(* Logix 5000 project; controller CIP vendor 1 type 14 code 106 rev 20.12; software revision 20.06; part 9 of 13 *)
(* tags used below, declared in another part *)
   MOA_OFF : DINT[10];
   MOA_ON : DINT[10];
   PV_Output_Status : INT[10];
   PV_Output_Status_IND : INT[10,16];
   PV_Status_Bit : BOOL;
(* MainProgram, continued *)

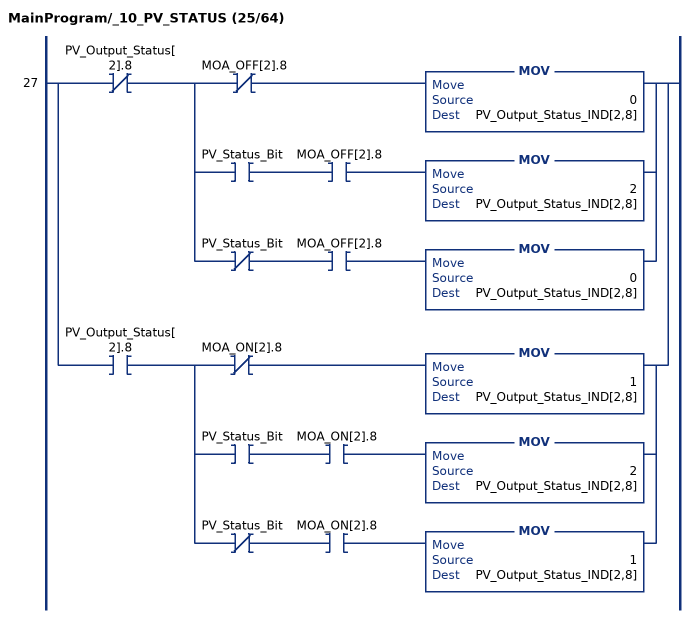
   [picture p157: MainProgram/_10_PV_STATUS rungs 27-27]
   27: [XIO(PV_Output_Status[2].8) [XIO(MOA_OFF[2].8) MOV(0,PV_Output_Status_IND[2,8]) ,XIC(PV_Status_Bit) XIC(MOA_OFF[2].8) MOV(2,PV_Output_Status_IND[2,8]) ,XIO(PV_Status_Bit) XIC(MOA_OFF[2].8) MOV(0,PV_Output_Status_IND[2,8]) ] ,XIC(PV_Output_Status[2].8) [XIO(MOA_ON[2].8) MOV(1,PV_Output_Status_IND[2,8]) ,XIC(PV_Status_Bit) XIC(MOA_ON[2].8) MOV(2,PV_Output_Status_IND[2,8]) ,XIO(PV_Status_Bit) XIC(MOA_ON[2].8) MOV(1,PV_Output_Status_IND[2,8]) ] ];
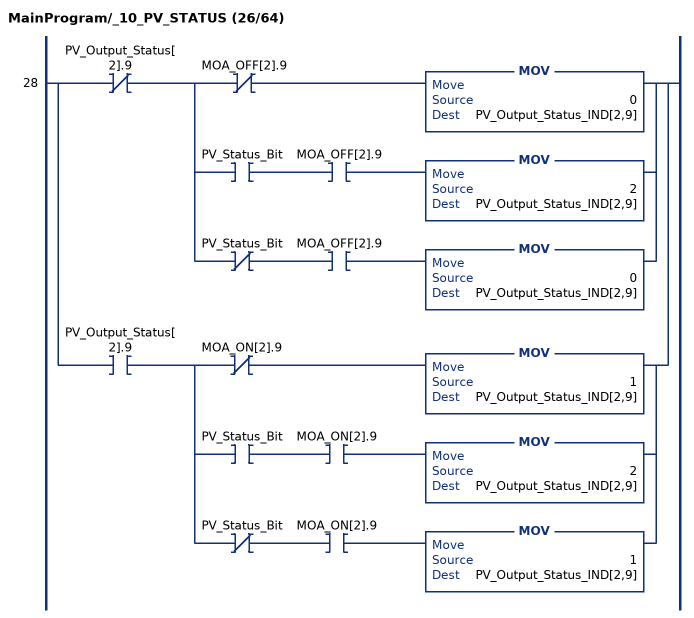
   28: [XIO(PV_Output_Status[2].9) [XIO(MOA_OFF[2].9) MOV(0,PV_Output_Status_IND[2,9]) ,XIC(PV_Status_Bit) XIC(MOA_OFF[2].9) MOV(2,PV_Output_Status_IND[2,9]) ,XIO(PV_Status_Bit) XIC(MOA_OFF[2].9) MOV(0,PV_Output_Status_IND[2,9]) ] ,XIC(PV_Output_Status[2].9) [XIO(MOA_ON[2].9) MOV(1,PV_Output_Status_IND[2,9]) ,XIC(PV_Status_Bit) XIC(MOA_ON[2].9) MOV(2,PV_Output_Status_IND[2,9]) ,XIO(PV_Status_Bit) XIC(MOA_ON[2].9) MOV(1,PV_Output_Status_IND[2,9]) ] ];
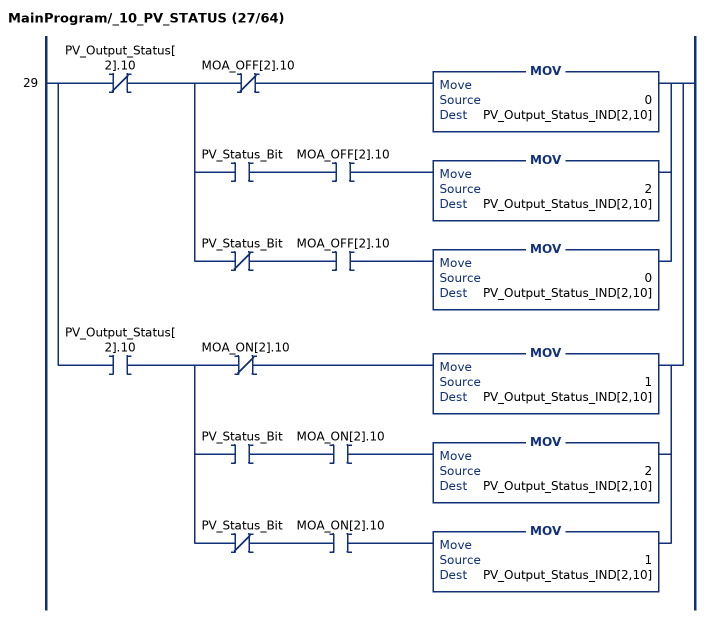
   29: [XIO(PV_Output_Status[2].10) [XIO(MOA_OFF[2].10) MOV(0,PV_Output_Status_IND[2,10]) ,XIC(PV_Status_Bit) XIC(MOA_OFF[2].10) MOV(2,PV_Output_Status_IND[2,10]) ,XIO(PV_Status_Bit) XIC(MOA_OFF[2].10) MOV(0,PV_Output_Status_IND[2,10]) ] ,XIC(PV_Output_Status[2].10) [XIO(MOA_ON[2].10) MOV(1,PV_Output_Status_IND[2,10]) ,XIC(PV_Status_Bit) XIC(MOA_ON[2].10) MOV(2,PV_Output_Status_IND[2,10]) ,XIO(PV_Status_Bit) XIC(MOA_ON[2].10) MOV(1,PV_Output_Status_IND[2,10]) ] ];
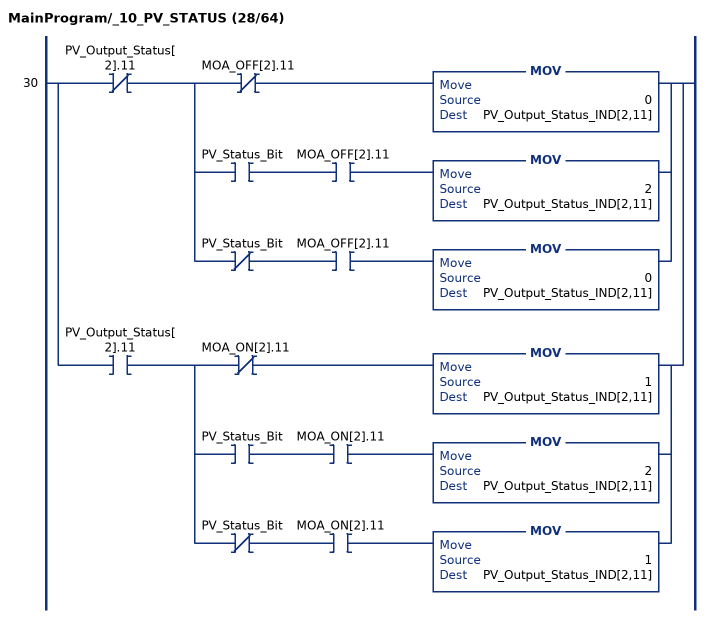
   30: [XIO(PV_Output_Status[2].11) [XIO(MOA_OFF[2].11) MOV(0,PV_Output_Status_IND[2,11]) ,XIC(PV_Status_Bit) XIC(MOA_OFF[2].11) MOV(2,PV_Output_Status_IND[2,11]) ,XIO(PV_Status_Bit) XIC(MOA_OFF[2].11) MOV(0,PV_Output_Status_IND[2,11]) ] ,XIC(PV_Output_Status[2].11) [XIO(MOA_ON[2].11) MOV(1,PV_Output_Status_IND[2,11]) ,XIC(PV_Status_Bit) XIC(MOA_ON[2].11) MOV(2,PV_Output_Status_IND[2,11]) ,XIO(PV_Status_Bit) XIC(MOA_ON[2].11) MOV(1,PV_Output_Status_IND[2,11]) ] ];
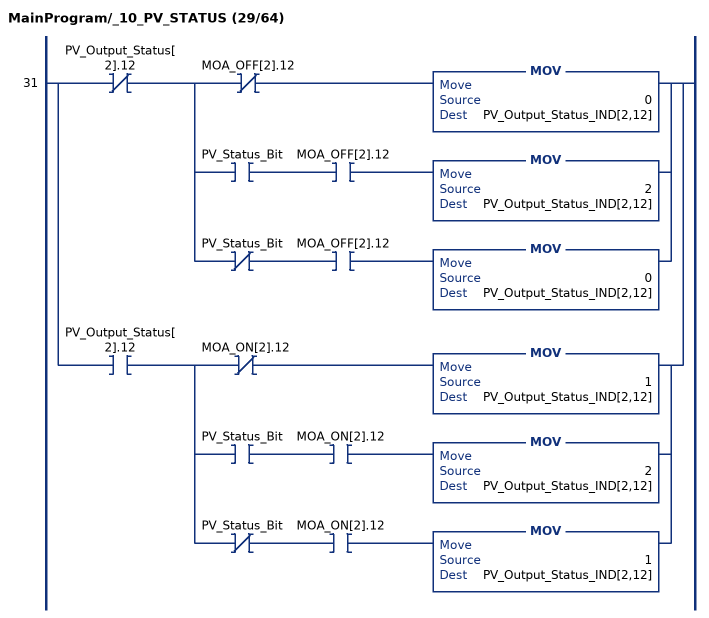
   31: [XIO(PV_Output_Status[2].12) [XIO(MOA_OFF[2].12) MOV(0,PV_Output_Status_IND[2,12]) ,XIC(PV_Status_Bit) XIC(MOA_OFF[2].12) MOV(2,PV_Output_Status_IND[2,12]) ,XIO(PV_Status_Bit) XIC(MOA_OFF[2].12) MOV(0,PV_Output_Status_IND[2,12]) ] ,XIC(PV_Output_Status[2].12) [XIO(MOA_ON[2].12) MOV(1,PV_Output_Status_IND[2,12]) ,XIC(PV_Status_Bit) XIC(MOA_ON[2].12) MOV(2,PV_Output_Status_IND[2,12]) ,XIO(PV_Status_Bit) XIC(MOA_ON[2].12) MOV(1,PV_Output_Status_IND[2,12]) ] ];
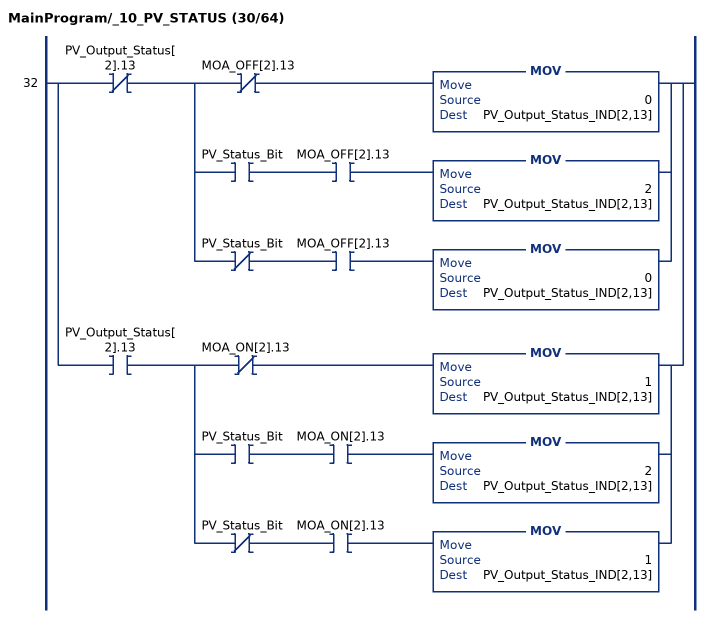
   32: [XIO(PV_Output_Status[2].13) [XIO(MOA_OFF[2].13) MOV(0,PV_Output_Status_IND[2,13]) ,XIC(PV_Status_Bit) XIC(MOA_OFF[2].13) MOV(2,PV_Output_Status_IND[2,13]) ,XIO(PV_Status_Bit) XIC(MOA_OFF[2].13) MOV(0,PV_Output_Status_IND[2,13]) ] ,XIC(PV_Output_Status[2].13) [XIO(MOA_ON[2].13) MOV(1,PV_Output_Status_IND[2,13]) ,XIC(PV_Status_Bit) XIC(MOA_ON[2].13) MOV(2,PV_Output_Status_IND[2,13]) ,XIO(PV_Status_Bit) XIC(MOA_ON[2].13) MOV(1,PV_Output_Status_IND[2,13]) ] ];
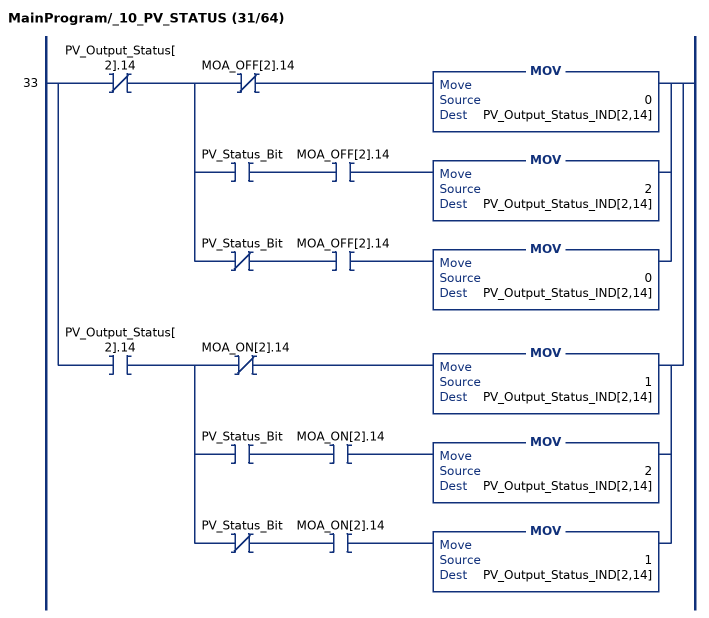
   33: [XIO(PV_Output_Status[2].14) [XIO(MOA_OFF[2].14) MOV(0,PV_Output_Status_IND[2,14]) ,XIC(PV_Status_Bit) XIC(MOA_OFF[2].14) MOV(2,PV_Output_Status_IND[2,14]) ,XIO(PV_Status_Bit) XIC(MOA_OFF[2].14) MOV(0,PV_Output_Status_IND[2,14]) ] ,XIC(PV_Output_Status[2].14) [XIO(MOA_ON[2].14) MOV(1,PV_Output_Status_IND[2,14]) ,XIC(PV_Status_Bit) XIC(MOA_ON[2].14) MOV(2,PV_Output_Status_IND[2,14]) ,XIO(PV_Status_Bit) XIC(MOA_ON[2].14) MOV(1,PV_Output_Status_IND[2,14]) ] ];
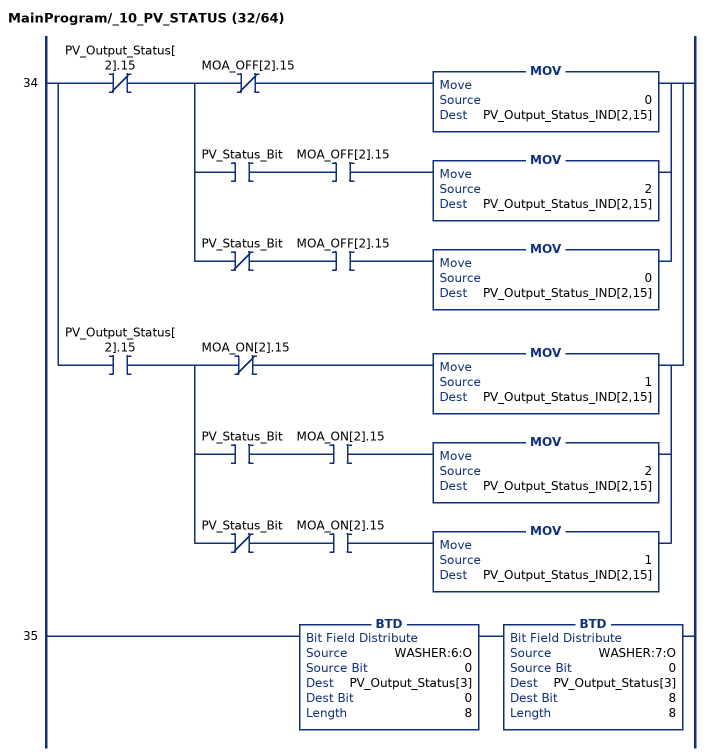
   34: [XIO(PV_Output_Status[2].15) [XIO(MOA_OFF[2].15) MOV(0,PV_Output_Status_IND[2,15]) ,XIC(PV_Status_Bit) XIC(MOA_OFF[2].15) MOV(2,PV_Output_Status_IND[2,15]) ,XIO(PV_Status_Bit) XIC(MOA_OFF[2].15) MOV(0,PV_Output_Status_IND[2,15]) ] ,XIC(PV_Output_Status[2].15) [XIO(MOA_ON[2].15) MOV(1,PV_Output_Status_IND[2,15]) ,XIC(PV_Status_Bit) XIC(MOA_ON[2].15) MOV(2,PV_Output_Status_IND[2,15]) ,XIO(PV_Status_Bit) XIC(MOA_ON[2].15) MOV(1,PV_Output_Status_IND[2,15]) ] ];
   35: BTD(WASHER:6:O,0,PV_Output_Status[3],0,8)BTD(WASHER:7:O,0,PV_Output_Status[3],8,8);
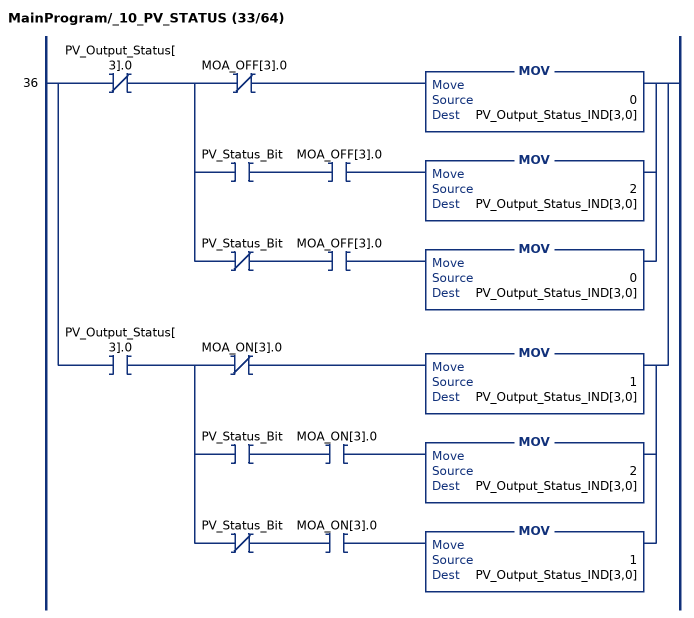
   36: [XIO(PV_Output_Status[3].0) [XIO(MOA_OFF[3].0) MOV(0,PV_Output_Status_IND[3,0]) ,XIC(PV_Status_Bit) XIC(MOA_OFF[3].0) MOV(2,PV_Output_Status_IND[3,0]) ,XIO(PV_Status_Bit) XIC(MOA_OFF[3].0) MOV(0,PV_Output_Status_IND[3,0]) ] ,XIC(PV_Output_Status[3].0) [XIO(MOA_ON[3].0) MOV(1,PV_Output_Status_IND[3,0]) ,XIC(PV_Status_Bit) XIC(MOA_ON[3].0) MOV(2,PV_Output_Status_IND[3,0]) ,XIO(PV_Status_Bit) XIC(MOA_ON[3].0) MOV(1,PV_Output_Status_IND[3,0]) ] ];
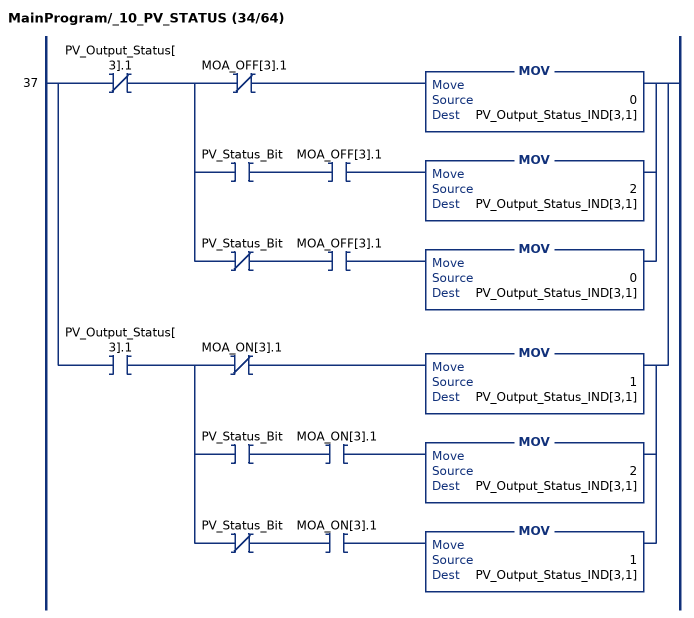
   37: [XIO(PV_Output_Status[3].1) [XIO(MOA_OFF[3].1) MOV(0,PV_Output_Status_IND[3,1]) ,XIC(PV_Status_Bit) XIC(MOA_OFF[3].1) MOV(2,PV_Output_Status_IND[3,1]) ,XIO(PV_Status_Bit) XIC(MOA_OFF[3].1) MOV(0,PV_Output_Status_IND[3,1]) ] ,XIC(PV_Output_Status[3].1) [XIO(MOA_ON[3].1) MOV(1,PV_Output_Status_IND[3,1]) ,XIC(PV_Status_Bit) XIC(MOA_ON[3].1) MOV(2,PV_Output_Status_IND[3,1]) ,XIO(PV_Status_Bit) XIC(MOA_ON[3].1) MOV(1,PV_Output_Status_IND[3,1]) ] ];
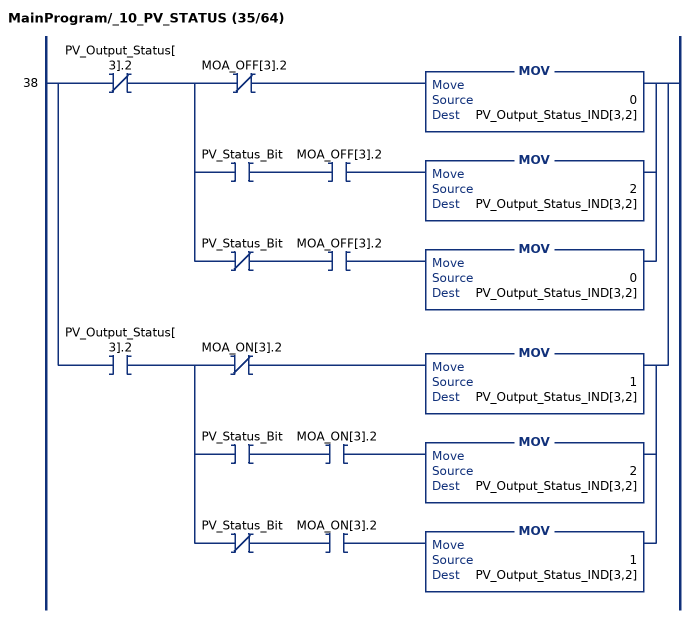
   38: [XIO(PV_Output_Status[3].2) [XIO(MOA_OFF[3].2) MOV(0,PV_Output_Status_IND[3,2]) ,XIC(PV_Status_Bit) XIC(MOA_OFF[3].2) MOV(2,PV_Output_Status_IND[3,2]) ,XIO(PV_Status_Bit) XIC(MOA_OFF[3].2) MOV(0,PV_Output_Status_IND[3,2]) ] ,XIC(PV_Output_Status[3].2) [XIO(MOA_ON[3].2) MOV(1,PV_Output_Status_IND[3,2]) ,XIC(PV_Status_Bit) XIC(MOA_ON[3].2) MOV(2,PV_Output_Status_IND[3,2]) ,XIO(PV_Status_Bit) XIC(MOA_ON[3].2) MOV(1,PV_Output_Status_IND[3,2]) ] ];
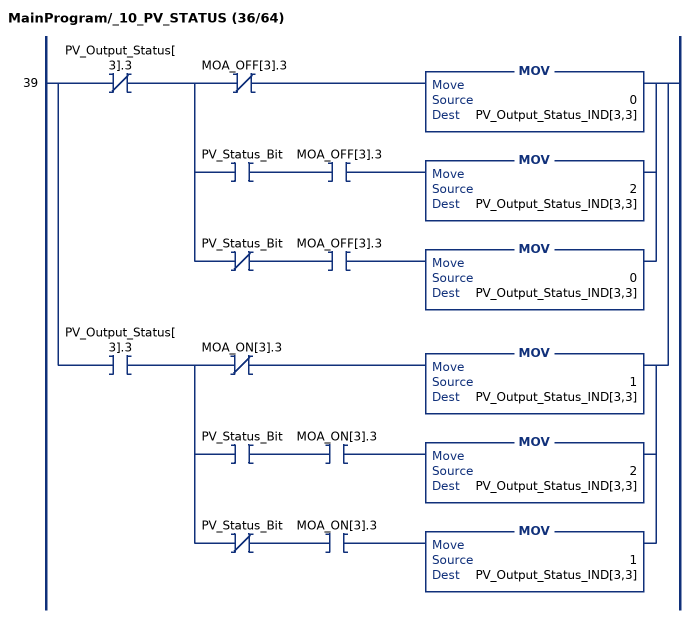
   39: [XIO(PV_Output_Status[3].3) [XIO(MOA_OFF[3].3) MOV(0,PV_Output_Status_IND[3,3]) ,XIC(PV_Status_Bit) XIC(MOA_OFF[3].3) MOV(2,PV_Output_Status_IND[3,3]) ,XIO(PV_Status_Bit) XIC(MOA_OFF[3].3) MOV(0,PV_Output_Status_IND[3,3]) ] ,XIC(PV_Output_Status[3].3) [XIO(MOA_ON[3].3) MOV(1,PV_Output_Status_IND[3,3]) ,XIC(PV_Status_Bit) XIC(MOA_ON[3].3) MOV(2,PV_Output_Status_IND[3,3]) ,XIO(PV_Status_Bit) XIC(MOA_ON[3].3) MOV(1,PV_Output_Status_IND[3,3]) ] ];
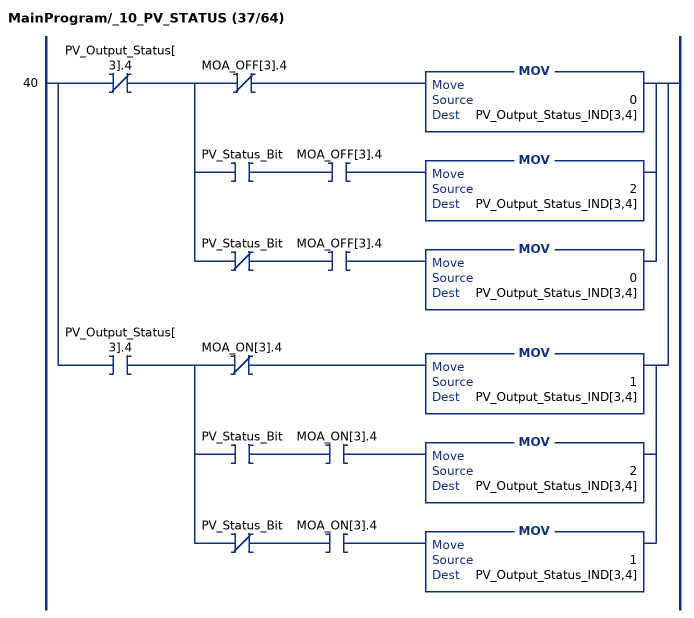
   40: [XIO(PV_Output_Status[3].4) [XIO(MOA_OFF[3].4) MOV(0,PV_Output_Status_IND[3,4]) ,XIC(PV_Status_Bit) XIC(MOA_OFF[3].4) MOV(2,PV_Output_Status_IND[3,4]) ,XIO(PV_Status_Bit) XIC(MOA_OFF[3].4) MOV(0,PV_Output_Status_IND[3,4]) ] ,XIC(PV_Output_Status[3].4) [XIO(MOA_ON[3].4) MOV(1,PV_Output_Status_IND[3,4]) ,XIC(PV_Status_Bit) XIC(MOA_ON[3].4) MOV(2,PV_Output_Status_IND[3,4]) ,XIO(PV_Status_Bit) XIC(MOA_ON[3].4) MOV(1,PV_Output_Status_IND[3,4]) ] ];
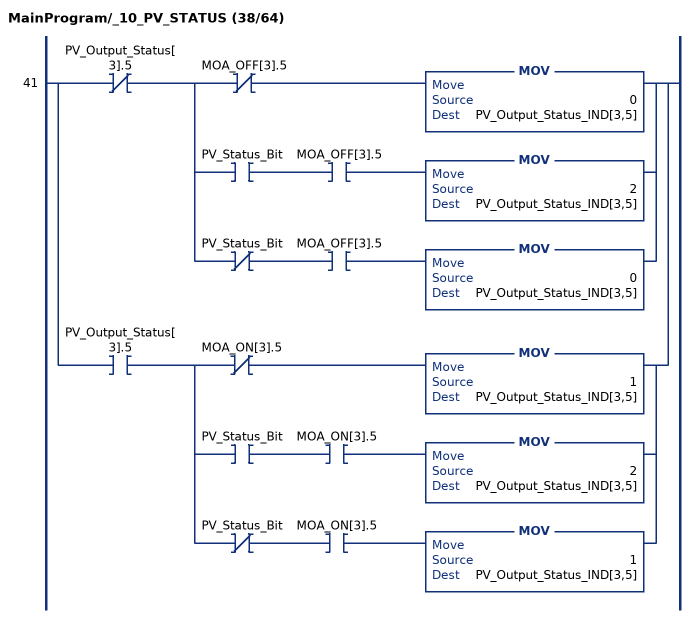
   41: [XIO(PV_Output_Status[3].5) [XIO(MOA_OFF[3].5) MOV(0,PV_Output_Status_IND[3,5]) ,XIC(PV_Status_Bit) XIC(MOA_OFF[3].5) MOV(2,PV_Output_Status_IND[3,5]) ,XIO(PV_Status_Bit) XIC(MOA_OFF[3].5) MOV(0,PV_Output_Status_IND[3,5]) ] ,XIC(PV_Output_Status[3].5) [XIO(MOA_ON[3].5) MOV(1,PV_Output_Status_IND[3,5]) ,XIC(PV_Status_Bit) XIC(MOA_ON[3].5) MOV(2,PV_Output_Status_IND[3,5]) ,XIO(PV_Status_Bit) XIC(MOA_ON[3].5) MOV(1,PV_Output_Status_IND[3,5]) ] ];
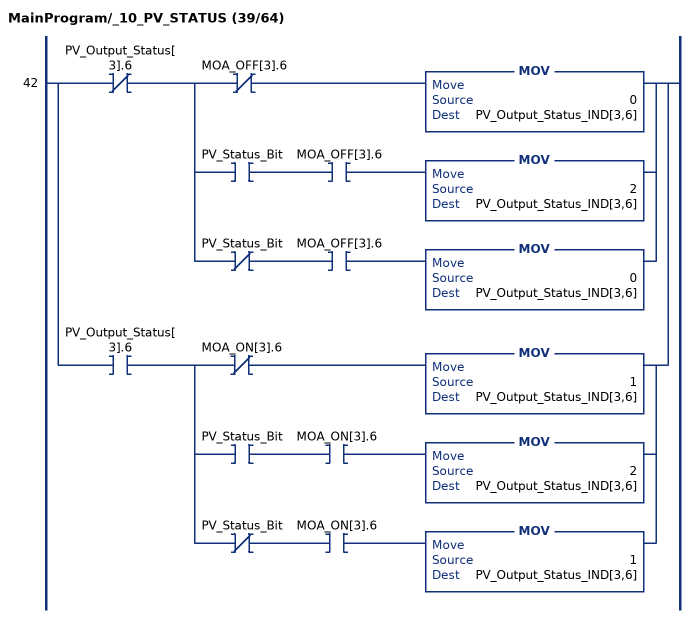
   42: [XIO(PV_Output_Status[3].6) [XIO(MOA_OFF[3].6) MOV(0,PV_Output_Status_IND[3,6]) ,XIC(PV_Status_Bit) XIC(MOA_OFF[3].6) MOV(2,PV_Output_Status_IND[3,6]) ,XIO(PV_Status_Bit) XIC(MOA_OFF[3].6) MOV(0,PV_Output_Status_IND[3,6]) ] ,XIC(PV_Output_Status[3].6) [XIO(MOA_ON[3].6) MOV(1,PV_Output_Status_IND[3,6]) ,XIC(PV_Status_Bit) XIC(MOA_ON[3].6) MOV(2,PV_Output_Status_IND[3,6]) ,XIO(PV_Status_Bit) XIC(MOA_ON[3].6) MOV(1,PV_Output_Status_IND[3,6]) ] ];
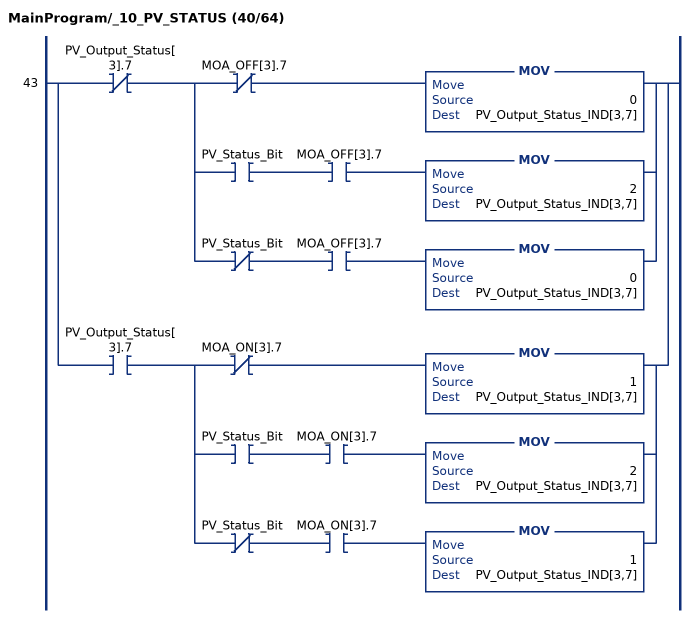
   43: [XIO(PV_Output_Status[3].7) [XIO(MOA_OFF[3].7) MOV(0,PV_Output_Status_IND[3,7]) ,XIC(PV_Status_Bit) XIC(MOA_OFF[3].7) MOV(2,PV_Output_Status_IND[3,7]) ,XIO(PV_Status_Bit) XIC(MOA_OFF[3].7) MOV(0,PV_Output_Status_IND[3,7]) ] ,XIC(PV_Output_Status[3].7) [XIO(MOA_ON[3].7) MOV(1,PV_Output_Status_IND[3,7]) ,XIC(PV_Status_Bit) XIC(MOA_ON[3].7) MOV(2,PV_Output_Status_IND[3,7]) ,XIO(PV_Status_Bit) XIC(MOA_ON[3].7) MOV(1,PV_Output_Status_IND[3,7]) ] ];
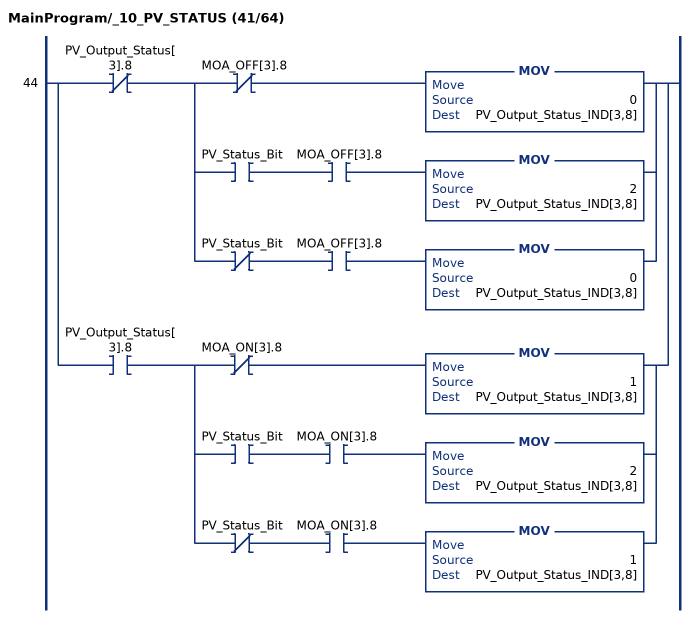
   44: [XIO(PV_Output_Status[3].8) [XIO(MOA_OFF[3].8) MOV(0,PV_Output_Status_IND[3,8]) ,XIC(PV_Status_Bit) XIC(MOA_OFF[3].8) MOV(2,PV_Output_Status_IND[3,8]) ,XIO(PV_Status_Bit) XIC(MOA_OFF[3].8) MOV(0,PV_Output_Status_IND[3,8]) ] ,XIC(PV_Output_Status[3].8) [XIO(MOA_ON[3].8) MOV(1,PV_Output_Status_IND[3,8]) ,XIC(PV_Status_Bit) XIC(MOA_ON[3].8) MOV(2,PV_Output_Status_IND[3,8]) ,XIO(PV_Status_Bit) XIC(MOA_ON[3].8) MOV(1,PV_Output_Status_IND[3,8]) ] ];
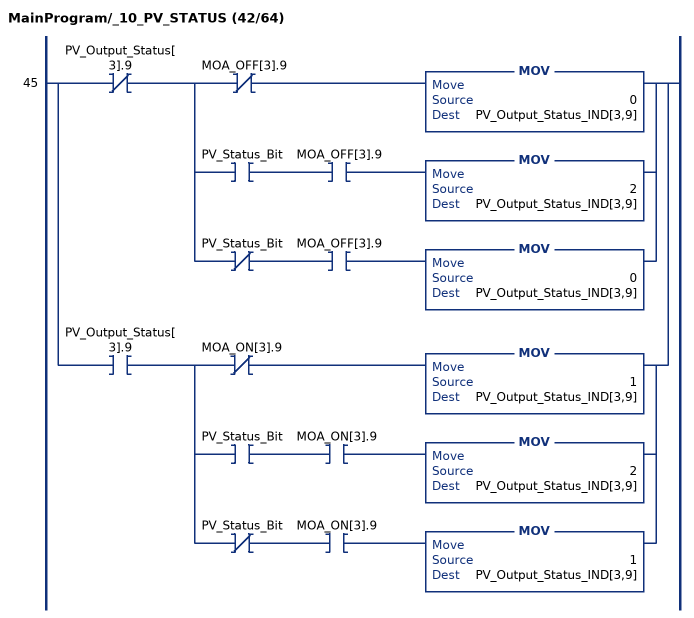
   45: [XIO(PV_Output_Status[3].9) [XIO(MOA_OFF[3].9) MOV(0,PV_Output_Status_IND[3,9]) ,XIC(PV_Status_Bit) XIC(MOA_OFF[3].9) MOV(2,PV_Output_Status_IND[3,9]) ,XIO(PV_Status_Bit) XIC(MOA_OFF[3].9) MOV(0,PV_Output_Status_IND[3,9]) ] ,XIC(PV_Output_Status[3].9) [XIO(MOA_ON[3].9) MOV(1,PV_Output_Status_IND[3,9]) ,XIC(PV_Status_Bit) XIC(MOA_ON[3].9) MOV(2,PV_Output_Status_IND[3,9]) ,XIO(PV_Status_Bit) XIC(MOA_ON[3].9) MOV(1,PV_Output_Status_IND[3,9]) ] ];
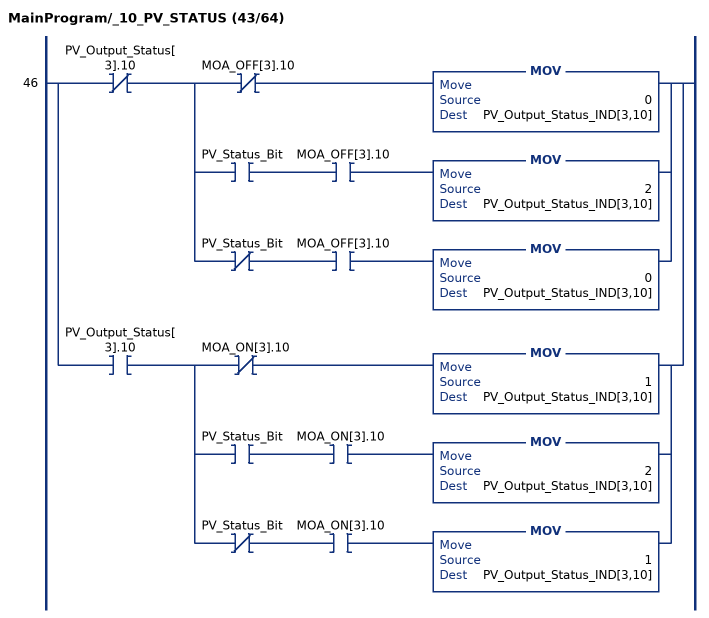
   46: [XIO(PV_Output_Status[3].10) [XIO(MOA_OFF[3].10) MOV(0,PV_Output_Status_IND[3,10]) ,XIC(PV_Status_Bit) XIC(MOA_OFF[3].10) MOV(2,PV_Output_Status_IND[3,10]) ,XIO(PV_Status_Bit) XIC(MOA_OFF[3].10) MOV(0,PV_Output_Status_IND[3,10]) ] ,XIC(PV_Output_Status[3].10) [XIO(MOA_ON[3].10) MOV(1,PV_Output_Status_IND[3,10]) ,XIC(PV_Status_Bit) XIC(MOA_ON[3].10) MOV(2,PV_Output_Status_IND[3,10]) ,XIO(PV_Status_Bit) XIC(MOA_ON[3].10) MOV(1,PV_Output_Status_IND[3,10]) ] ];
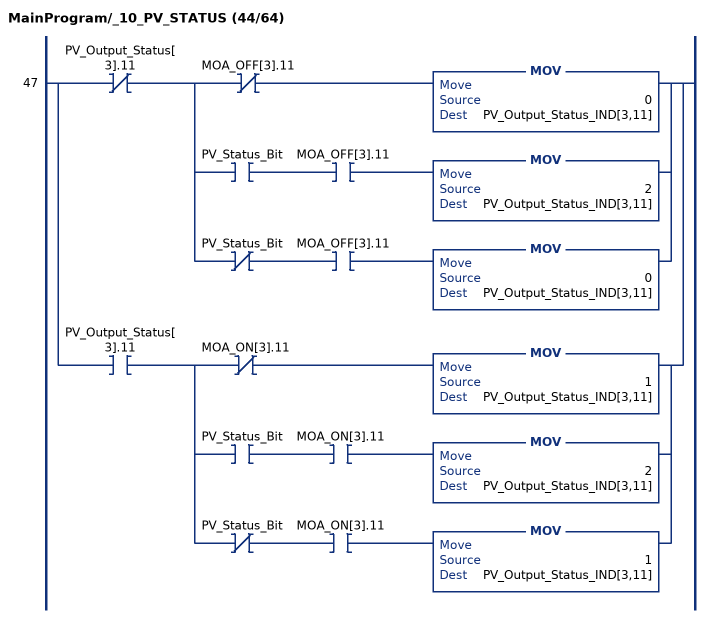
   47: [XIO(PV_Output_Status[3].11) [XIO(MOA_OFF[3].11) MOV(0,PV_Output_Status_IND[3,11]) ,XIC(PV_Status_Bit) XIC(MOA_OFF[3].11) MOV(2,PV_Output_Status_IND[3,11]) ,XIO(PV_Status_Bit) XIC(MOA_OFF[3].11) MOV(0,PV_Output_Status_IND[3,11]) ] ,XIC(PV_Output_Status[3].11) [XIO(MOA_ON[3].11) MOV(1,PV_Output_Status_IND[3,11]) ,XIC(PV_Status_Bit) XIC(MOA_ON[3].11) MOV(2,PV_Output_Status_IND[3,11]) ,XIO(PV_Status_Bit) XIC(MOA_ON[3].11) MOV(1,PV_Output_Status_IND[3,11]) ] ];
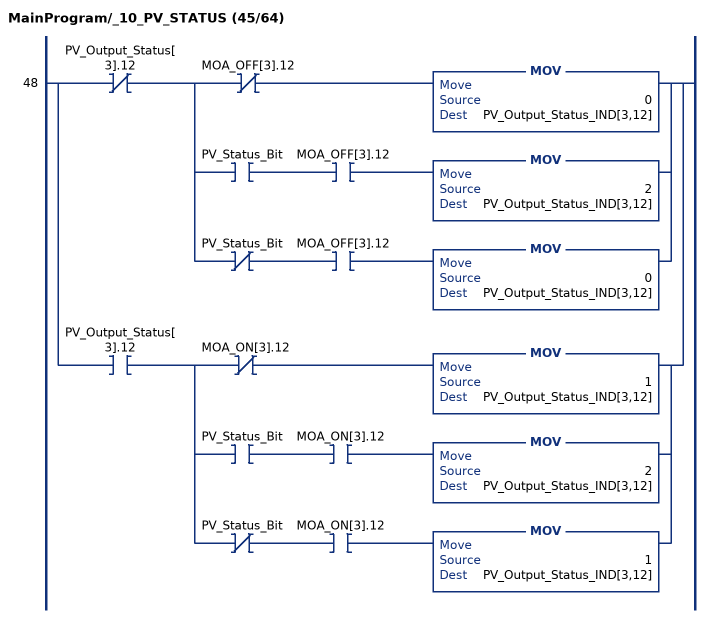
   48: [XIO(PV_Output_Status[3].12) [XIO(MOA_OFF[3].12) MOV(0,PV_Output_Status_IND[3,12]) ,XIC(PV_Status_Bit) XIC(MOA_OFF[3].12) MOV(2,PV_Output_Status_IND[3,12]) ,XIO(PV_Status_Bit) XIC(MOA_OFF[3].12) MOV(0,PV_Output_Status_IND[3,12]) ] ,XIC(PV_Output_Status[3].12) [XIO(MOA_ON[3].12) MOV(1,PV_Output_Status_IND[3,12]) ,XIC(PV_Status_Bit) XIC(MOA_ON[3].12) MOV(2,PV_Output_Status_IND[3,12]) ,XIO(PV_Status_Bit) XIC(MOA_ON[3].12) MOV(1,PV_Output_Status_IND[3,12]) ] ];
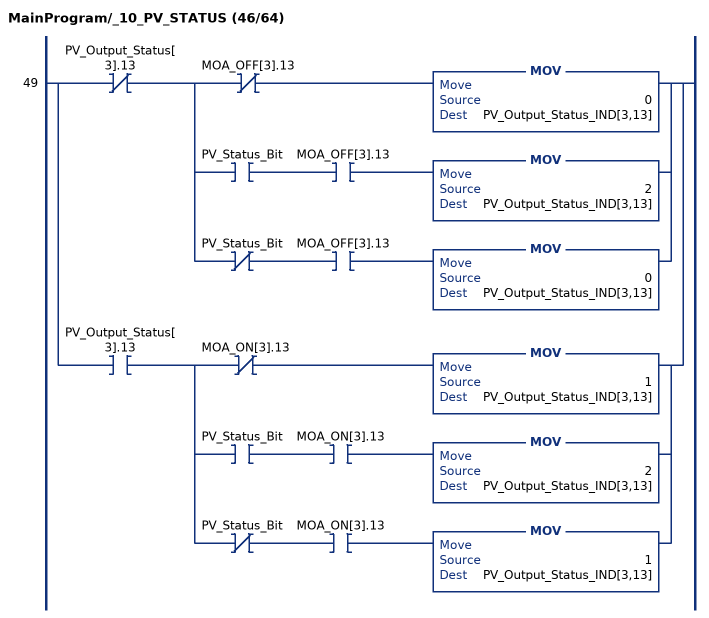
   49: [XIO(PV_Output_Status[3].13) [XIO(MOA_OFF[3].13) MOV(0,PV_Output_Status_IND[3,13]) ,XIC(PV_Status_Bit) XIC(MOA_OFF[3].13) MOV(2,PV_Output_Status_IND[3,13]) ,XIO(PV_Status_Bit) XIC(MOA_OFF[3].13) MOV(0,PV_Output_Status_IND[3,13]) ] ,XIC(PV_Output_Status[3].13) [XIO(MOA_ON[3].13) MOV(1,PV_Output_Status_IND[3,13]) ,XIC(PV_Status_Bit) XIC(MOA_ON[3].13) MOV(2,PV_Output_Status_IND[3,13]) ,XIO(PV_Status_Bit) XIC(MOA_ON[3].13) MOV(1,PV_Output_Status_IND[3,13]) ] ];
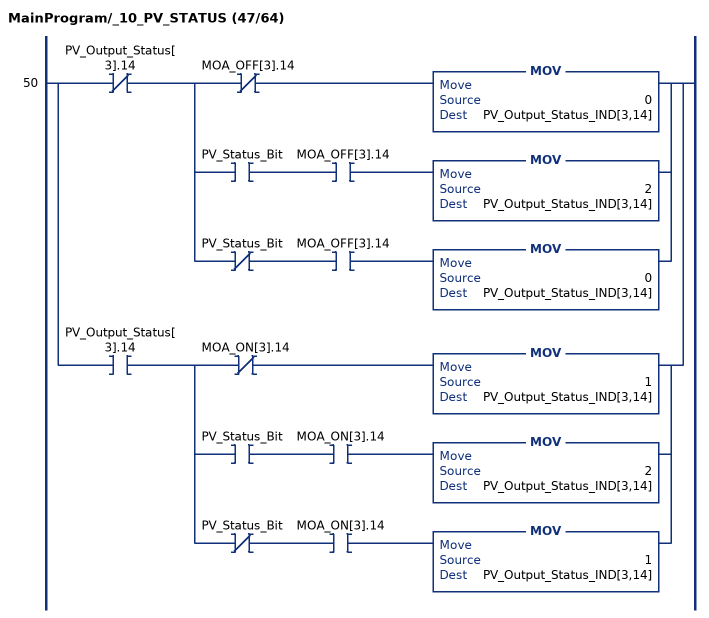
   50: [XIO(PV_Output_Status[3].14) [XIO(MOA_OFF[3].14) MOV(0,PV_Output_Status_IND[3,14]) ,XIC(PV_Status_Bit) XIC(MOA_OFF[3].14) MOV(2,PV_Output_Status_IND[3,14]) ,XIO(PV_Status_Bit) XIC(MOA_OFF[3].14) MOV(0,PV_Output_Status_IND[3,14]) ] ,XIC(PV_Output_Status[3].14) [XIO(MOA_ON[3].14) MOV(1,PV_Output_Status_IND[3,14]) ,XIC(PV_Status_Bit) XIC(MOA_ON[3].14) MOV(2,PV_Output_Status_IND[3,14]) ,XIO(PV_Status_Bit) XIC(MOA_ON[3].14) MOV(1,PV_Output_Status_IND[3,14]) ] ];
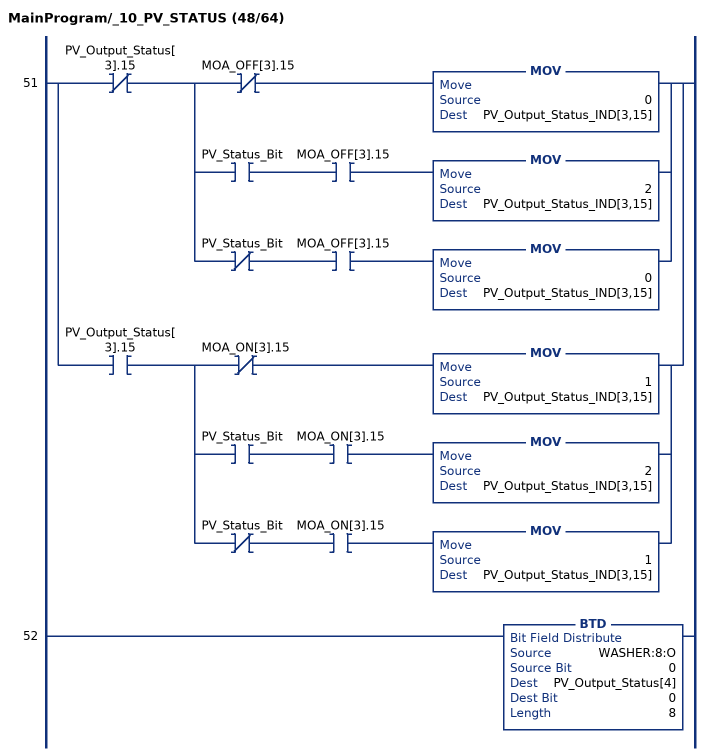
   51: [XIO(PV_Output_Status[3].15) [XIO(MOA_OFF[3].15) MOV(0,PV_Output_Status_IND[3,15]) ,XIC(PV_Status_Bit) XIC(MOA_OFF[3].15) MOV(2,PV_Output_Status_IND[3,15]) ,XIO(PV_Status_Bit) XIC(MOA_OFF[3].15) MOV(0,PV_Output_Status_IND[3,15]) ] ,XIC(PV_Output_Status[3].15) [XIO(MOA_ON[3].15) MOV(1,PV_Output_Status_IND[3,15]) ,XIC(PV_Status_Bit) XIC(MOA_ON[3].15) MOV(2,PV_Output_Status_IND[3,15]) ,XIO(PV_Status_Bit) XIC(MOA_ON[3].15) MOV(1,PV_Output_Status_IND[3,15]) ] ];
   52: BTD(WASHER:8:O,0,PV_Output_Status[4],0,8);
